FUNCTION_BLOCK AB_LAST_4 (* MERGE 4 AB in 1 AB (LAST WRITER WINS, generic FB) - welcher Socket zuletzt geschrieben hat, gewinnt und wird sofort an OUT durchgereicht *)
  (* Standard: 61499-2; Description: Copyright (c) 2026 Meisterschulen am Ostbahnhof This program and the accompanying materials are made available under the terms of the Eclipse Public License 2.0 which is available at https://www.eclipse.org/legal/epl-2.0/ SPDX-License-Identifier: EPL-2.0 *)
  (* Version 1.0, 2026-11-06, Franz Höpfinger, Meisterschulen am Ostbahnhof, generic FB GEN_AB_LAST (N Sockets), Verhalten in FORTE *)
  PACKAGE adapter::events::unidirectional;
  IMPORT eclipse4diac::core::GenericClassName;
  {SET_ATTRIBUTE(eclipse4diac::core::GenericClassName, 'GEN_AB_LAST')}
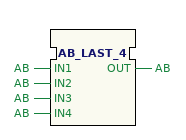
  SOCKETS
    IN1 : adapter::types::unidirectional::AB;
    IN2 : adapter::types::unidirectional::AB;
    IN3 : adapter::types::unidirectional::AB;
    IN4 : adapter::types::unidirectional::AB;
  END_SOCKETS
  PLUGS
    OUT : adapter::types::unidirectional::AB;
  END_PLUGS
END_FUNCTION_BLOCK
